(* Logix 5000 project; controller ProductSortingConveyor vendor 1 type 14 code 164 rev 37.11; software revision 37.00 *)

TASK MainTask (continuous, watchdog 500 ms) : MainProgram

MODULES
   Local : vendor 1 type 14 code 164 (ICP 0, rev 37.11)
END_MODULES

VAR_GLOBAL   (* controller tags *)
   Blue_Button : BOOL;
   Blue_Load : BOOL;
   Box_Present : BOOL;
   CollisionSensor_Blue : BOOL;
   CollisionSensor_Green : BOOL;
   CollisionSensor_Orange : BOOL;
   CollisionSensor_Purple : BOOL;
   CollisionSensor_Red : BOOL;
   CollisionSensor_Yellow : BOOL;
   Conveyor : BOOL;
   Cycle_Done : BOOL;
   Detect_Trigger : BOOL;
   Distance : REAL;
   Green_Button : BOOL;
   Green_Load : BOOL;
   OneShot : BOOL;
   Orange_Button : BOOL;
   Orange_Load : BOOL;
   Plunger_Blue : BOOL;
   Plunger_Green : BOOL;
   Plunger_Orange : BOOL;
   Plunger_Purple : BOOL;
   Plunger_Red : BOOL;
   Plunger_Timer : TIMER := (PRE := 500);
   Plunger_Yellow : BOOL;
   Purple_Button : BOOL;
   Purple_Load : BOOL;
   Red_Button : BOOL;
   Red_Load : BOOL;
   Start_Button : BOOL;
   Stop_Button : BOOL;
   Stopper_Blue : BOOL;
   Stopper_Blue_Cmd : BOOL;
   Stopper_Green : BOOL;
   Stopper_Green_Cmd : BOOL;
   Stopper_Orange : BOOL;
   Stopper_Orange_Cmd : BOOL;
   Stopper_Purple : BOOL;
   Stopper_Purple_Cmd : BOOL;
   Stopper_Red : BOOL;
   Stopper_Red_Cmd : BOOL;
   Stopper_Yellow : BOOL;
   Stopper_Yellow_Cmd : BOOL;
   Timer_Blue : TIMER := (PRE := 300);
   Timer_Green : TIMER := (PRE := 300);
   Timer_Orange : TIMER := (PRE := 300);
   Timer_Purple : TIMER := (PRE := 300);
   Timer_Red : TIMER := (PRE := 300);
   Timer_Yellow : TIMER := (PRE := 300);
   Yellow_Button : BOOL;
   Yellow_Load : BOOL;
END_VAR

PROGRAM MainProgram   (* main routine MainRoutine *)
VAR
   BoxType : DINT;
END_VAR

ROUTINE MainRoutine   (* ladder *)
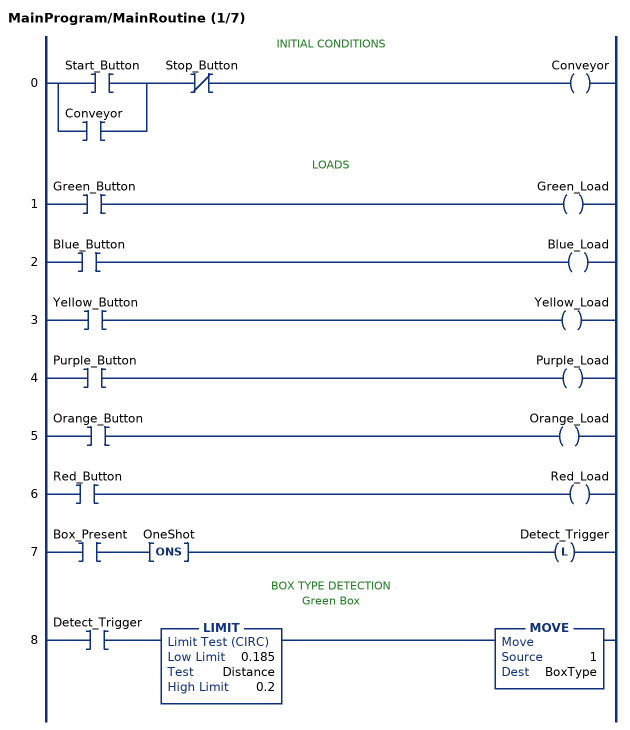
   // INITIAL CONDITIONS
   0: [XIC(Start_Button) ,XIC(Conveyor) ]XIO(Stop_Button)OTE(Conveyor);
   // LOADS
   1: XIC(Green_Button)OTE(Green_Load);
   2: XIC(Blue_Button)OTE(Blue_Load);
   3: XIC(Yellow_Button)OTE(Yellow_Load);
   4: XIC(Purple_Button)OTE(Purple_Load);
   5: XIC(Orange_Button)OTE(Orange_Load);
   6: XIC(Red_Button)OTE(Red_Load);
   7: XIC(Box_Present)ONS(OneShot)OTL(Detect_Trigger);
   // BOX TYPE DETECTION
   // Green Box
   8: XIC(Detect_Trigger)LIMIT(0.185,Distance,0.2)MOVE(1,BoxType);
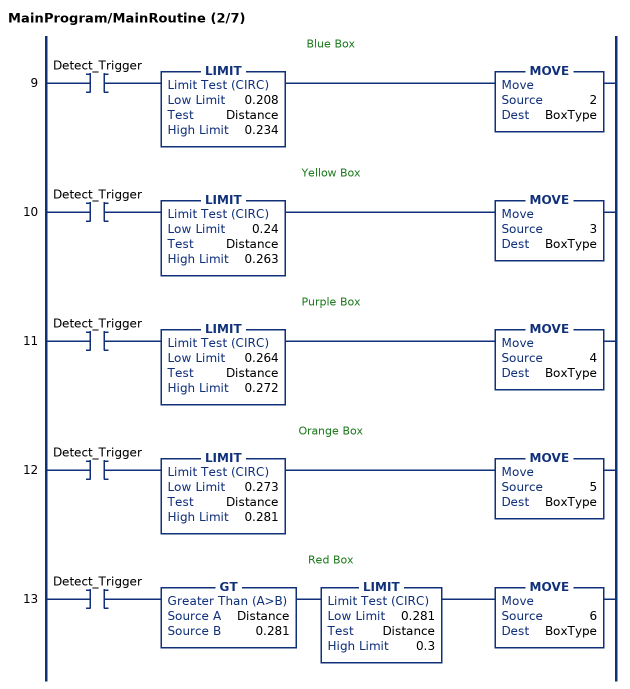
   // Blue Box
   9: XIC(Detect_Trigger)LIMIT(0.208,Distance,0.234)MOVE(2,BoxType);
   // Yellow Box
   10: XIC(Detect_Trigger)LIMIT(0.24,Distance,0.263)MOVE(3,BoxType);
   // Purple Box
   11: XIC(Detect_Trigger)LIMIT(0.264,Distance,0.272)MOVE(4,BoxType);
   // Orange Box
   12: XIC(Detect_Trigger)LIMIT(0.273,Distance,0.281)MOVE(5,BoxType);
   // Red Box
   13: XIC(Detect_Trigger)GT(Distance,0.281)LIMIT(0.281,Distance,0.3)MOVE(6,BoxType);
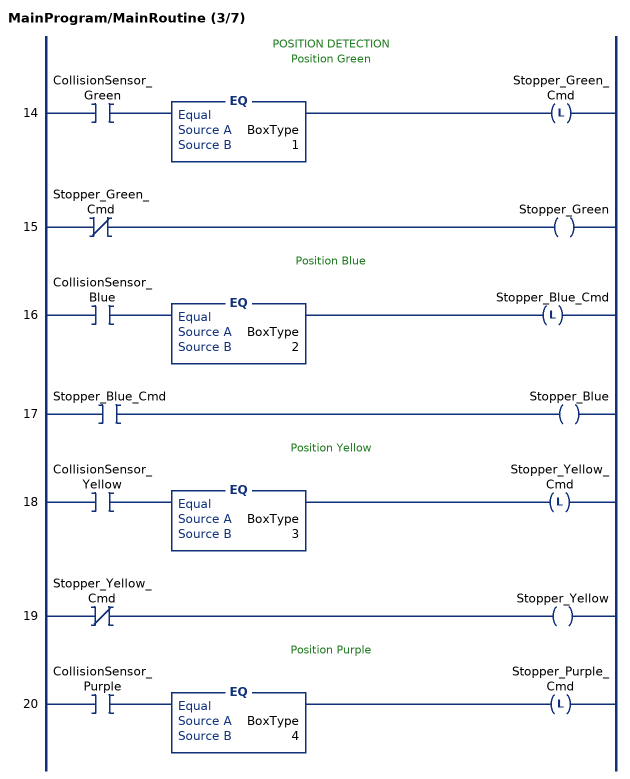
   // POSITION DETECTION
   // Position Green
   14: XIC(CollisionSensor_Green)EQ(BoxType,1)OTL(Stopper_Green_Cmd);
   15: XIO(Stopper_Green_Cmd)OTE(Stopper_Green);
   // Position Blue
   16: XIC(CollisionSensor_Blue)EQ(BoxType,2)OTL(Stopper_Blue_Cmd);
   17: XIC(Stopper_Blue_Cmd)OTE(Stopper_Blue);
   // Position Yellow
   18: XIC(CollisionSensor_Yellow)EQ(BoxType,3)OTL(Stopper_Yellow_Cmd);
   19: XIO(Stopper_Yellow_Cmd)OTE(Stopper_Yellow);
   // Position Purple
   20: XIC(CollisionSensor_Purple)EQ(BoxType,4)OTL(Stopper_Purple_Cmd);
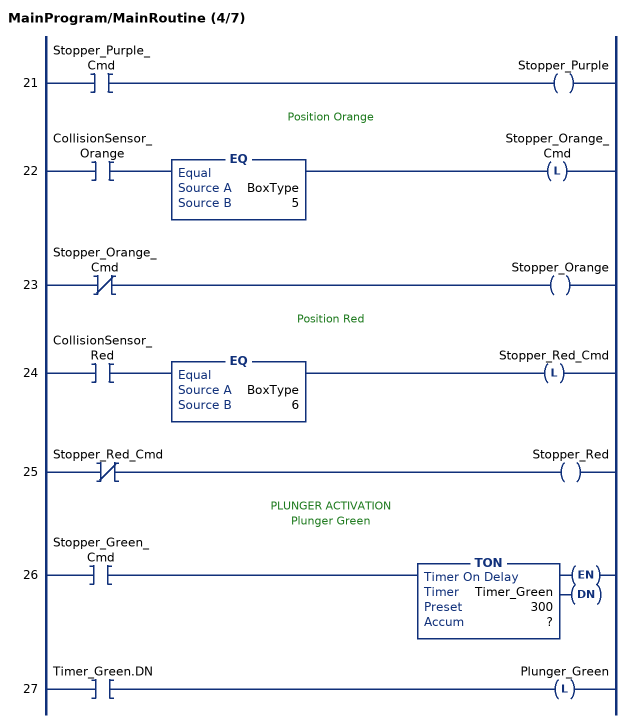
   21: XIC(Stopper_Purple_Cmd)OTE(Stopper_Purple);
   // Position Orange
   22: XIC(CollisionSensor_Orange)EQ(BoxType,5)OTL(Stopper_Orange_Cmd);
   23: XIO(Stopper_Orange_Cmd)OTE(Stopper_Orange);
   // Position Red
   24: XIC(CollisionSensor_Red)EQ(BoxType,6)OTL(Stopper_Red_Cmd);
   25: XIO(Stopper_Red_Cmd)OTE(Stopper_Red);
   // PLUNGER ACTIVATION
   // Plunger Green
   26: XIC(Stopper_Green_Cmd)TON(Timer_Green,?,?);
   27: XIC(Timer_Green.DN)OTL(Plunger_Green);
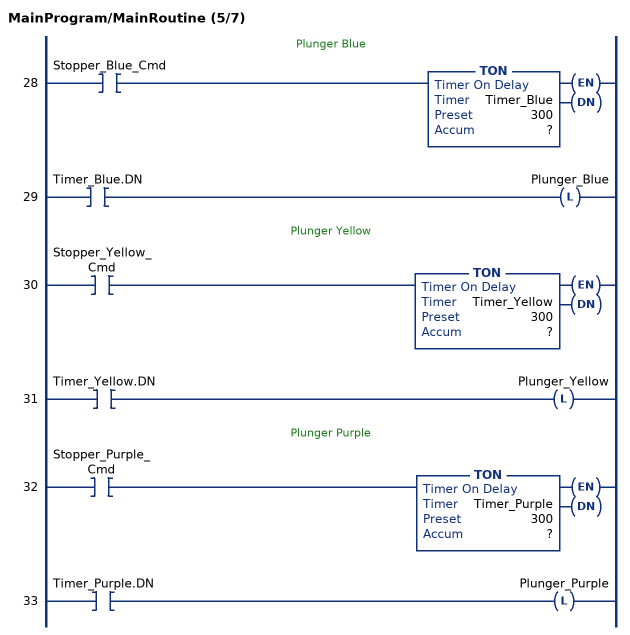
   // Plunger Blue
   28: XIC(Stopper_Blue_Cmd)TON(Timer_Blue,?,?);
   29: XIC(Timer_Blue.DN)OTL(Plunger_Blue);
   // Plunger Yellow
   30: XIC(Stopper_Yellow_Cmd)TON(Timer_Yellow,?,?);
   31: XIC(Timer_Yellow.DN)OTL(Plunger_Yellow);
   // Plunger Purple
   32: XIC(Stopper_Purple_Cmd)TON(Timer_Purple,?,?);
   33: XIC(Timer_Purple.DN)OTL(Plunger_Purple);
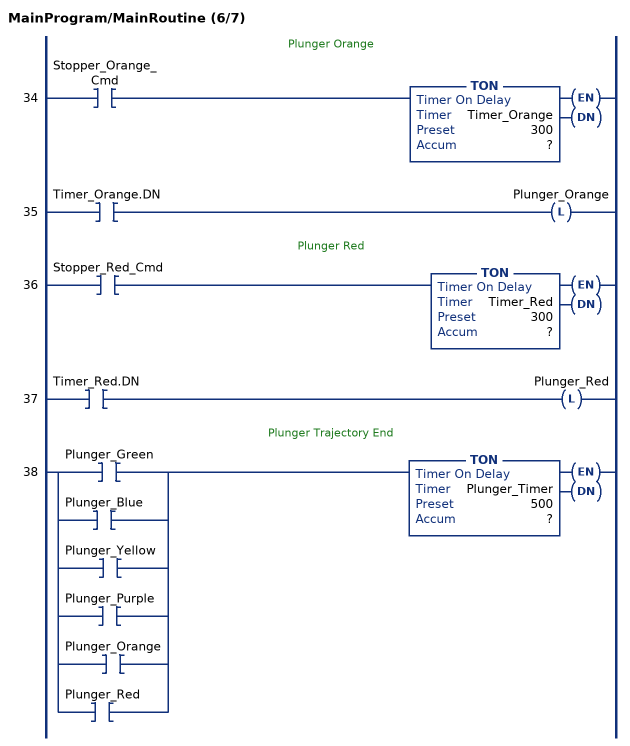
   // Plunger Orange
   34: XIC(Stopper_Orange_Cmd)TON(Timer_Orange,?,?);
   35: XIC(Timer_Orange.DN)OTL(Plunger_Orange);
   // Plunger Red
   36: XIC(Stopper_Red_Cmd)TON(Timer_Red,?,?);
   37: XIC(Timer_Red.DN)OTL(Plunger_Red);
   // Plunger Trajectory End
   38: [XIC(Plunger_Green) ,XIC(Plunger_Blue) ,XIC(Plunger_Yellow) ,XIC(Plunger_Purple) ,XIC(Plunger_Orange) ,XIC(Plunger_Red) ]TON(Plunger_Timer,?,?);
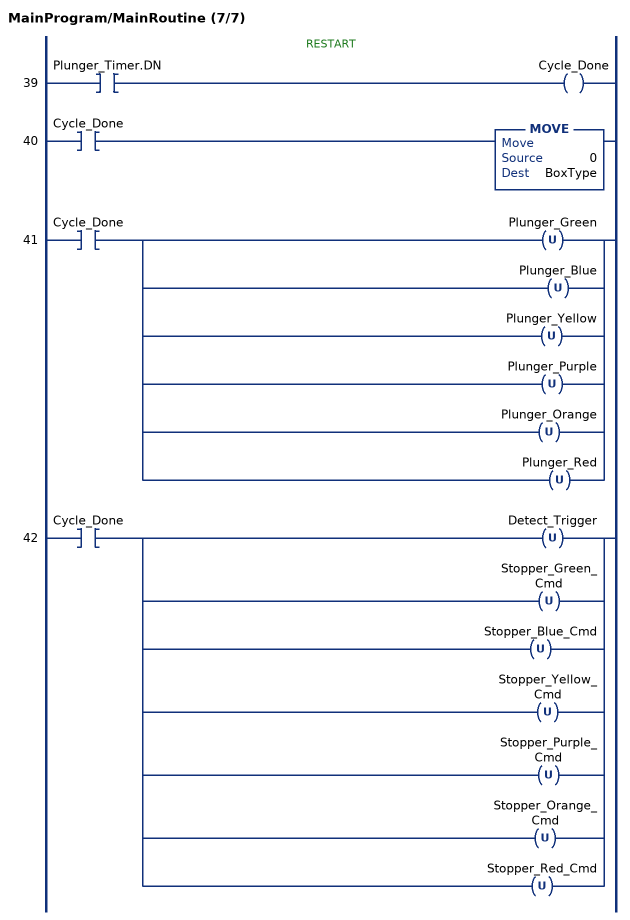
   // RESTART
   39: XIC(Plunger_Timer.DN)OTE(Cycle_Done);
   40: XIC(Cycle_Done)MOVE(0,BoxType);
   41: XIC(Cycle_Done)[OTU(Plunger_Green) ,OTU(Plunger_Blue) ,OTU(Plunger_Yellow) ,OTU(Plunger_Purple) ,OTU(Plunger_Orange) ,OTU(Plunger_Red) ];
   42: XIC(Cycle_Done)[OTU(Detect_Trigger) ,OTU(Stopper_Green_Cmd) ,OTU(Stopper_Blue_Cmd) ,OTU(Stopper_Yellow_Cmd) ,OTU(Stopper_Purple_Cmd) ,OTU(Stopper_Orange_Cmd) ,OTU(Stopper_Red_Cmd) ];
END_ROUTINE
END_PROGRAM
